ACTION ACT_ResetDrives:
// =============================================================
// ACT_ResetDrives
// Kasowanie bledow wszystkich falownikow
// =============================================================
//
// Dziala na ZBOCZE bitu xCmdResetDrives. Blok napedu wystawia
// impuls 200 ms na bicie 7 ControlWord - falownik NORD kasuje
// blad zboczem, nie poziomem.
//
// Kasujemy WSZYSTKIE napedy, takze te zablokowane w
// axDriveEnabled: skasowanie bledu niczego nie uruchamia,
// a chcemy widziec czysty obraz maszyny.
//
// Bit zdejmujemy sami, zeby nie trzeba bylo tego robic recznie
// w podgladzie online.

// -------------------------------------------------------------
// KASOWANIE RECZNE - bitem
// -------------------------------------------------------------

rtrgResetDrv(CLK := xCmdResetDrives);

IF rtrgResetDrv.Q THEN

	FOR i := 1 TO cNumDrives DO
		fbNord[i].M_Reset();
	END_FOR

	xCmdResetDrives	:= FALSE;
	xResetFailed	:= FALSE;

END_IF


// -------------------------------------------------------------
// KASOWANIE AUTOMATYCZNE - po wcisnieciu START
// -------------------------------------------------------------
//
// Kasujemy tylko te napedy, ktore faktycznie zglaszaja blad,
// i tylko ograniczona liczbe razy. Bez tego limitu maszyna
// dobijalaby sie w nieskonczonosc do napedu, ktory ma realny
// powod stac - a to wygladaloby jak "nic sie nie dzieje".

IF NOT xResetInProgress THEN
	RETURN;
END_IF


// Czysto - konczymy
IF NOT xAnyDriveFault THEN
	xResetInProgress	:= FALSE;
	nResetTries			:= 0;
	tonResetGap(IN := FALSE);
	RETURN;
END_IF


// Proby wyczerpane - dalej decyduje czlowiek
IF nResetTries >= cResetTries THEN
	xResetInProgress	:= FALSE;
	xResetFailed		:= TRUE;
	tonResetGap(IN := FALSE);
	RETURN;
END_IF


// Pierwsza proba od razu, kolejne co tResetGap
IF nResetTries = 0 THEN
	xDoResetPulse := TRUE;
ELSE
	tonResetGap(IN := TRUE, PT := tResetGap);
	xDoResetPulse := tonResetGap.Q;
END_IF

IF NOT xDoResetPulse THEN
	RETURN;
END_IF

tonResetGap(IN := FALSE);


FOR i := 1 TO cNumDrives DO
	IF axDrvFault[i] THEN
		fbNord[i].M_Reset();
	END_IF
END_FOR

nResetTries := nResetTries + 1;
END_ACTION

ACTION ACT_Sequence:
// =============================================================
// ACT_Sequence
// Wirtualna paleta idaca trasa maszyny
// =============================================================
//
// Paleta ZATRZYMUJE SIE na kazdej stacji. Cykl wyglada tak:
//
//   przejazd  para transporterow pracuje przez tStepTime,
//             potem OBA staja
//   praca     transportery stoja, dziala mechanika stacji
//             (kazdy ruch silownika przez tCylTime)
//   i dalej
//
// Czujnikow nie ma, wiec o zakonczeniu kazdej fazy decyduje
// czas. Po dolozeniu czujnikow te czasowki zastapi warunek
// "paleta na pozycji" i "silownik w polozeniu".
//
// TRASA:
//   poz. 1..11   dobre:   1-2-3-4-5-6-7-8-11-12-13
//   poz. 12..16  odrzut:  8-10-14-15-16  (8 -> 10 lancuchem)
//
// Przydzial falownikow do stacji:
//   st.1  -> 8     st.5  -> 5     st.9  -> 7      st.13 -> 15
//   st.2  -> 9     st.6  -> 6     st.10 -> 16     st.14 -> 17
//   st.3  -> 10    st.7  -> 11    st.11 -> 13     st.15 -> 18
//   st.4  -> 4     st.8  -> 12    st.12 -> 14     st.16 -> 19


// Zadanie ruchu kasujemy w kazdym cyklu - faza ustawia je od nowa
FOR i := 1 TO 20 DO
	axRunReq[i] := FALSE;
END_FOR

tThisStep := tCylTime;


// -------------------------------------------------------------
// START I STOP
// -------------------------------------------------------------

rtrgStart(CLK := START_TEST);

IF rtrgStart.Q THEN

	nIdx	:= 0;			// najpierw sprowadzamy mechanike
	nSub	:= 0;
	xMoving	:= FALSE;
	tonStep(IN := FALSE);

	xResetFailed := FALSE;
	nResetTries  := 0;
	tonResetGap(IN := FALSE);

	IF xAutoResetOnStart AND xAnyDriveFault THEN
		xResetInProgress := TRUE;
	END_IF

END_IF


IF NOT START_TEST THEN
	tonStep(IN := FALSE);
	sPhase := 'STOP - START_TEST = FALSE';
	ACT_ClearCoils();
	RETURN;
END_IF


IF NOT xSafetyOK THEN
	tonStep(IN := FALSE);
	sPhase := 'STOP - brak zezwolenia bezpieczenstwa';
	RETURN;
END_IF


IF xResetInProgress THEN
	tonStep(IN := FALSE);
	sPhase := CONCAT('kasowanie bledow falownikow - proba ',
	                 INT_TO_STRING(nResetTries));
	RETURN;
END_IF


// -------------------------------------------------------------
// TRYB RECZNY POJEDYNCZEGO SILOWNIKA
// -------------------------------------------------------------
//
// Ma pierwszenstwo przed sekwencja - transportery stoja,
// bo axRunReq zostalo wykasowane na gorze.

IF nManCyl <> 0 THEN
	ACT_ManualCyl();
	tonStep(IN := FALSE);
	RETURN;
END_IF


// -------------------------------------------------------------
// ZMIANA KROKU
// -------------------------------------------------------------
//
// Kazdy krok dostaje czasowke od zera i wlasne uzbrojenie
// czujnika. Bez tego krok dziedziczylby resztke po poprzednim.

xNewStep := (nIdx <> nIdxOld) OR (nSub <> nSubOld) OR (xMoving <> xMovingOld);

nIdxOld		:= nIdx;
nSubOld		:= nSub;
xMovingOld	:= xMoving;

IF xNewStep THEN
	tonStep(IN := FALSE);
	xStepArmed   := FALSE;
	xStepTimeout := FALSE;
END_IF


// Krok sam zglosi, na co czeka. Kasujemy co cykl.
xWaitSensor := FALSE;
xSensorOK   := FALSE;


// -------------------------------------------------------------
// FAZA
// -------------------------------------------------------------

IF xMoving THEN
	ACT_Move();
ELSE
	ACT_Work();
END_IF


// -------------------------------------------------------------
// KONIEC KROKU: CZUJNIK ALBO WATCHDOG
// -------------------------------------------------------------
//
// Krok czujnikowy konczy sie czujnikiem. Czasowka pracuje wtedy
// tylko jako watchdog - jesli to ONA zdecyduje, zapala sie
// xStepTimeout i wiadomo, ze czujnik nie przyszedl.
//
// Czujnik musi byc najpierw WOLNY (xStepArmed). Inaczej krok
// zaliczylby stan sprzed przejazdu albo czujnik zwarty na stale.

IF xUseSensors AND xWaitSensor THEN
	tThisStep := tMoveTimeout;
END_IF

tonStep(IN := TRUE, PT := tThisStep);
xAdvance := tonStep.Q;

// Watchdog wylaczony - czasowka nie ma prawa zakonczyc kroku
// czujnikowego. Krok stoi, dopoki nie przyjdzie sam czujnik.
IF xUseSensors AND xWaitSensor AND NOT xStepWatchdog THEN
	xAdvance := FALSE;
END_IF

IF xUseSensors AND xWaitSensor AND xAdvance THEN
	xStepTimeout := TRUE;
	nTimeouts    := nTimeouts + 1;
END_IF

IF NOT xSensorOK THEN
	xStepArmed := TRUE;
END_IF

IF xUseSensors AND xWaitSensor AND xStepArmed AND xSensorOK THEN
	xAdvance := TRUE;
END_IF

IF xAdvance THEN
	tonStep(IN := FALSE);
END_IF
END_ACTION

ACTION ACT_TestFeed:
// =============================================================
// ACT_TestFeed
// Proba calosciowa: st.1 -> desztaplarka -> stacja 4
// =============================================================
//
// Waska sciezka transportu na czas proby. NIE korzysta z tabeli
// trasy w ACT_Sequence - wozi tylko tam, gdzie trzeba:
//
//   1. dowozi stos ze stacji 1 na stacje 3 (czujnik IN2),
//   2. czeka, az desztaplarka zwolni palete,
//   3. wywozi ja przez stacje 4 robiac test dociskow,
//   4. ZATRZYMUJE ja na koncu stacji 4 - do recznego zabrania.
//
// Napedy: st.1 -> 8, st.2 -> 9, st.3 -> 10, st.4 -> 4.
// Rolki dociskowe (falownik 3) zostaja wylaczone.
//
// Cewki dociskow przepisujemy CO CYKL - ACT_ClearCoils zeruje
// je przy zdjetym START_TEST, wiec krok, ktory ich nie odswieza,
// stracilby sterowanie zaworem.


xFeedNewStep := (nFeedStep <> nFeedStepOld);
nFeedStepOld := nFeedStep;

IF xFeedNewStep THEN
	tonFeedStep(IN := FALSE);
	xFeedArmed := FALSE;
END_IF

tonFeedStep(IN := TRUE, PT := tFeedStep);
xFeedAdvance := tonFeedStep.Q AND NOT xFeedNewStep;


// Tor B ma WLASNA czasowke i wlasne uzbrojenie czujnika -
// inaczej dwie palety deptalyby sobie po jednym liczniku.
//
// UWAGA NA ZBOCZE KROKU MIEDZY TORAMI.
// Flagi xOutNewStep / xOutAdvance sa liczone TU, na poczatku
// akcji. Jesli inny tor wpisze torowi B numer kroku PO tym
// miejscu, krok wykona sie jeszcze w tym samym cyklu - ze stara
// flaga xOutAdvance, odziedziczona po kroku 0, gdzie czasowka
// dawno wybila. Krok przeskoczylby natychmiast.
//
// Wlasnie tak ginal przejazd ze stacji 5 na 6: krok 180 trwal
// JEDEN CYKL zadania, naped 5 dostawal zadanie na 10 ms i tor
// szedl dalej, jakby paleta juz przejechala.
//
// Dlatego zaden tor nie wpisuje numeru kroku innemu torowi.
// Zglasza tylko zadanie (xOutStart), a tor podnosi je SAM,
// w swoim kroku 0 - i wtedy pierwszy cykl nowego kroku jest
// juz zwyklym zboczem, z wyzerowana czasowka.

xOutNewStep := (nOutStep <> nOutStepOld);
nOutStepOld := nOutStep;

IF xOutNewStep THEN
	tonOutStep(IN := FALSE);
	xOutArmed := FALSE;
END_IF

tonOutStep(IN := TRUE, PT := tOutStep);
xOutAdvance := tonOutStep.Q AND NOT xOutNewStep;


xOut2NewStep := (nOut2Step <> nOut2StepOld);
nOut2StepOld := nOut2Step;

IF xOut2NewStep THEN
	tonOut2Step(IN := FALSE);
	xOut2Armed := FALSE;
END_IF

tonOut2Step(IN := TRUE, PT := tOut2Step);
xOut2Advance := tonOut2Step.Q AND NOT xOut2NewStep;


xOut3NewStep := (nOut3Step <> nOut3StepOld);
nOut3StepOld := nOut3Step;

IF xOut3NewStep THEN
	tonOut3Step(IN := FALSE);
	xOut3Armed := FALSE;
END_IF

tonOut3Step(IN := TRUE, PT := tOut3Step);
xOut3Advance := tonOut3Step.Q AND NOT xOut3NewStep;


// Czas pchania palety do blokady stacji 5 - liczony od wejscia
// w krok 80, niezalezny od czasowki kroku.
tonSt05Push(IN := (nFeedStep = 80), PT := tSt05_Push);

// Ile blokada stacji 5 stoi juz OPUSZCZONA. Nie ma na niej
// czujnika, wiec liczymy od zdjecia komendy wysuwu - tyle, ile
// dajemy kazdemu silownikowi na dojscie do polozenia.
tonSt05BlockDown(IN := NOT xFeed05_Block, PT := tCylTime);

// Od IN7 na stacji 8 do opuszczenia rolek pod paleta NOK.
// Liczona OSOBNO od tFeedSt08Stop - to sa dwie rozne rzeczy,
// wiec MOGA byc w dowolnej kolejnosci i dowolnie dalekie.
//
// Odliczamy od FLAGI OBECNOSCI, a nie od numeru kroku. Krok 215
// trwa tylko tFeedSt08Stop; przy dluzszym tSt08_DropDelay timer
// nie zdazyl dobiec do konca i zerowal sie przy przejsciu do
// kroku 218. Rolki nie schodzily wcale, a to, ze pierwsza paleta
// wygladala dobrze, robil krok 220 toru B3 - i tylko wtedy, gdy
// lancuch byl akurat wolny.
tonSt08Drop(IN := xSt08_AtStation, PT := tSt08_DropDelay);


rtrgFeedStart(CLK := START_FEED);

IF rtrgFeedStart.Q THEN
	nFeedStep  := 0;

	// Tor B tez od zera - inaczej po ponownym starcie dokanczal
	// by trase palety, ktorej juz tam nie ma.
	nOutStep   := 0;
	nOut2Step  := 0;
	nOut3Step  := 0;
	xSt05_Done := FALSE;
	xOutStart  := FALSE;
	xOut2Start := FALSE;
	xOut3Start := FALSE;
	xSt08_RollDown  := FALSE;
	xSt08_AtStation := FALSE;
END_IF


// Falowniki po zatrzymaniu runtime'u zglaszaja blad komunikacji
// i same z niego nie wyjda. Kasujemy go przy starcie, tak samo
// jak robi to START_TEST - inaczej za kazdym razem trzeba by
// pamietac o xCmdResetDrives.
IF rtrgFeedStart.Q AND xAutoResetOnStart AND xAnyDriveFault THEN
	xResetInProgress := TRUE;
	nResetTries      := 0;
	xResetFailed     := FALSE;
END_IF


// Domyslnie: cala mechanika w polozeniu spoczynkowym.
// Krok, ktory czegos potrzebuje, podaje to sam.
xFeedPressOn   := FALSE;
xFeedPressLoOn := FALSE;
xFeed05_Block  := FALSE;
xFeed05_Lift   := FALSE;
xFeed05_Jaws   := FALSE;
xFeed05_Pull   := FALSE;
tFeedStep      := tSt04_EntryToPress;
tOutStep       := tCylTime;
tOut2Step      := tCylTime;
tOut3Step      := tCylTime;

// Rolki domyslnie W GORZE - transport wzdluz. Tylko przejazd
// lancuchem opuszcza je swiadomie.
xFeedRoll08Up  := TRUE;
xFeedRoll10Up  := TRUE;


IF NOT START_FEED THEN
	sFeedPhase := 'DOWOZ - stop, START_FEED = FALSE';
END_IF


IF START_FEED AND xSafetyOK THEN

	CASE nFeedStep OF

	0:
		sFeedPhase := 'DOWOZ 0 czekam na potwierdzenie palet na st.1';

		// Bit SAM sie zdejmuje po przyjeciu. Dzieki temu po
		// oproznieniu stosu maszyna nie rusza w pustke, tylko
		// czeka na kolejne potwierdzenie operatora.
		//
		// Jesli IN2 juz widzi stos, to on STOI na stacji 3
		// i nie ma czego dowozic - idziemy od razu do pracy
		// desztaplarki. "Juz u celu" nie jest powodem do
		// czekania.
		IF xSt01_StackReady AND NOT xPal_St03 THEN
			xSt01_StackReady := FALSE;
			nFeedStep        := 10;
		END_IF

		IF xSt01_StackReady AND xPal_St03 THEN
			sFeedPhase       := 'DOWOZ 0 stos JUZ na st.3 - pomijam dowoz';
			xSt01_StackReady := FALSE;
			nFeedStep        := 20;
		END_IF

	10:
		sFeedPhase := 'DOWOZ 1 stos jedzie st.1 -> st.3, czekam na IN2';
		axRunReq[8]  := TRUE;
		axRunReq[9]  := TRUE;
		axRunReq[10] := TRUE;

		IF NOT xPal_St03 THEN xFeedArmed := TRUE; END_IF

		IF xPal_St03 AND NOT xFeedArmed THEN
			sFeedPhase := 'DOWOZ 1 IN2 JUZ zaslonony - odslon i zaslon ponownie';
		END_IF

		IF xFeedArmed AND xPal_St03 THEN nFeedStep := 15; END_IF

	15:
		// Dobieg po czujniku - stos dojezdza pod szczeki.
		// Przy tFeedSt03Stop = 0 krok trwa jeden cykl zadania.
		sFeedPhase := 'DOWOZ 1b dobieg stosu po IN2';
		axRunReq[9]  := TRUE;
		axRunReq[10] := TRUE;
		tFeedStep    := tFeedSt03Stop;

		IF xFeedAdvance THEN nFeedStep := 20; END_IF

	20:
		// Transportery STOJA - desztaplarka pracuje na stosie.
		sFeedPhase := 'DOWOZ 2 stos na st.3 - czekam na zwolnienie palety';

		IF xDe_PalletReleased THEN nFeedStep := 30; END_IF

	30:
		sFeedPhase := 'DOWOZ 3 paleta jedzie na st.4, czekam na IN3';

		// Paleta zaslaniajaca JUZ czujnik konca stacji 4 minela
		// wjazd pod rolki. Czekanie na IN3 bylo by czekaniem na
		// zdarzenie, ktore sie nie powtorzy - jedziemy dalej.
		IF xFeedNewStep AND xPal_St04End THEN
			sFeedPhase := 'DOWOZ 3 paleta JUZ na koncu st.4 - pomijam docisk';
			nFeedStep  := 75;
		END_IF

		axRunReq[10] := TRUE;
		axRunReq[4]  := TRUE;

		IF NOT xPal_St04In THEN xFeedArmed := TRUE; END_IF

		IF xPal_St04In AND NOT xFeedArmed THEN
			sFeedPhase := 'DOWOZ 3 IN3 JUZ zaslonony - odslon i zaslon ponownie';
		END_IF

		IF xFeedArmed AND xPal_St04In THEN nFeedStep := 40; END_IF

	40:
		sFeedPhase := 'ST.4 wjazd pod rolki - odstep przed dociskiem';
		axRunReq[10] := TRUE;
		axRunReq[4]  := TRUE;
		axRunReq[3]  := TRUE;   // rolki dociskowe
		tFeedStep    := tSt04_EntryToPress;

		IF xFeedAdvance THEN nFeedStep := 50; END_IF

	50:
		sFeedPhase := 'ST.4 dociski gorne schodza na deski';
		axRunReq[10] := TRUE;
		axRunReq[4]  := TRUE;
		axRunReq[3]  := TRUE;   // rolki dociskowe
		xFeedPressOn := TRUE;
		tFeedStep    := tSt04_UpToLo;

		IF xFeedAdvance THEN nFeedStep := 60; END_IF

	60:
		sFeedPhase := 'ST.4 TEST - czekam na koniec testu (IN4)';
		axRunReq[10]   := TRUE;
		axRunReq[4]    := TRUE;
		axRunReq[3]  := TRUE;   // rolki dociskowe
		xFeedPressOn   := TRUE;
		xFeedPressLoOn := TRUE;

		IF NOT xPal_St04End THEN xFeedArmed := TRUE; END_IF

		IF xPal_St04End AND NOT xFeedArmed THEN
			sFeedPhase := 'ST.4 IN4 JUZ zaslonony - odslon i zaslon ponownie';
		END_IF

		IF xFeedArmed AND xPal_St04End THEN nFeedStep := 70; END_IF

	70:
		// Dociski juz cofniete - kroki wyzej ich nie podaja.
		sFeedPhase := 'ST.4 koniec testu - dociski cofniete, dojazd';
		axRunReq[4] := TRUE;
		tFeedStep   := tSt04_StopDelay;

		IF xFeedAdvance THEN nFeedStep := 75; END_IF

	75:
		// BRAMKA MIEDZY TORAMI. Stacja 5 to zasob wspolny:
		// jej transporter i blokada obsluguja raz palete
		// wyjezdzajaca, raz wjezdzajaca. Wjazd moze ruszyc
		// dopiero wtedy, gdy poprzednia paleta zjechala ze
		// stacji 5 - czyli tor B jest wolny (0) albo minal
		// juz przejazd na stacje 6 (>= 200).
		//
		// Paleta czeka na koncu stacji 4, napedy stoja.
		sFeedPhase := 'ST.4 koniec - czekam, az zwolni sie stacja 5';

		IF (nOutStep = 0) OR (nOutStep >= 200) THEN
			nFeedStep := 80;
		END_IF

	80:
		// Blokada wysuwa sie RAZEM z ruszeniem palety ze stacji 4.
		// To ona zatrzymuje palete na stacji 5 - nie ma tam
		// czujnika, wiec musi czekac na palete, a nie odwrotnie.
		// Napedy pracuja TYLKO przez tSt05_Push, a nie przez caly
		// krok. Paleta opiera sie o blokade po kilku sekundach
		// i od tej chwili transporter mieli pod stojaca paleta -
		// tak przeciazylismy naped 5. Reszta kroku to juz tylko
		// uspokojenie palety, z zatrzymanymi napedami.
		sFeedPhase := 'ST.4 -> ST.5 przejazd, blokada juz wysunieta';
		xFeed05_Block := TRUE;
		tFeedStep   := tFeedToSt05;

		IF NOT tonSt05Push.Q THEN
			axRunReq[4] := TRUE;
			axRunReq[5] := TRUE;
		END_IF

		IF tonSt05Push.Q THEN
			sFeedPhase := 'ST.5 paleta na blokadzie - napedy staja';
		END_IF

		IF xFeedAdvance THEN nFeedStep := 100; END_IF


	// -----------------------------------------------------
	// STACJA 5 - TEST ROZRYWANIA
	// -----------------------------------------------------
	//
	// Transportery STOJA. Kolejnosc wg zalozen: blokada,
	// podniesienie szczek, chwyt, szesc silownikow rozrywajacych
	// w gore i w dol, zwolnienie, opuszczenie blokady.
	//
	// Kazdy krok podaje SWOJ pelny stan cewek - przepisujemy je
	// na dole akcji, w kazdym cyklu.

	100:
		// Paleta oparla sie o blokade. Transportery juz stoja,
		// dajemy jej uspokoic sie, zanim ruszy mechanika.
		sFeedPhase := 'ST.5 1/8 paleta na blokadzie - uspokojenie';
		xFeed05_Block := TRUE;
		tFeedStep     := tSt05_Settle;
		IF xFeedAdvance THEN nFeedStep := 110; END_IF

	110:
		sFeedPhase := 'ST.5 2/8 szczeki ida w gore';
		xFeed05_Block := TRUE;
		xFeed05_Lift  := TRUE;
		tFeedStep     := tCylTime;
		IF xFeedAdvance THEN nFeedStep := 120; END_IF

	120:
		sFeedPhase := 'ST.5 3/8 szczeki zamykaja sie na deskach';
		xFeed05_Block := TRUE;
		xFeed05_Lift  := TRUE;
		xFeed05_Jaws  := TRUE;
		tFeedStep     := tCylTime;
		IF xFeedAdvance THEN nFeedStep := 130; END_IF

	130:
		sFeedPhase := 'ST.5 4/8 ROZRYWANIE - silowniki ida w gore';
		xFeed05_Block := TRUE;
		xFeed05_Lift  := TRUE;
		xFeed05_Jaws  := TRUE;
		xFeed05_Pull  := TRUE;
		tFeedStep     := tCylTime;
		IF xFeedAdvance THEN nFeedStep := 140; END_IF

	140:
		sFeedPhase := 'ST.5 5/8 silowniki rozrywajace ida w dol';
		xFeed05_Block := TRUE;
		xFeed05_Lift  := TRUE;
		xFeed05_Jaws  := TRUE;
		tFeedStep     := tCylTime;
		IF xFeedAdvance THEN nFeedStep := 150; END_IF

	150:
		sFeedPhase := 'ST.5 6/8 szczeki otwieraja sie';
		xFeed05_Block := TRUE;
		xFeed05_Lift  := TRUE;
		tFeedStep     := tCylTime;
		IF xFeedAdvance THEN nFeedStep := 160; END_IF

	160:
		sFeedPhase := 'ST.5 7/8 szczeki ida w dol';
		xFeed05_Block := TRUE;
		tFeedStep     := tCylTime;
		IF xFeedAdvance THEN nFeedStep := 170; END_IF

	170:
		// PRZEKAZANIE PALETY TOROWI B.
		//
		// Tu konczy sie zadanie toru A. Paleta ma wolna droge
		// (blokada opuszczona) i od tej chwili jedzie na stacje
		// 16 SAMA, sekwencja nOutStep. Tor A wraca po nastepna.
		//
		// xSt05_Done to sygnal dla desztaplarki - na nim wydaje
		// kolejna palete, nie czekajac na stacje 16.
		//
		// Jesli tor B jeszcze pracuje, paleta czeka tutaj:
		// stoi na stacji 5 z opuszczona blokada, napedy staja.
		sFeedPhase := 'ST.5 8/8 blokada opuszcza sie';
		tFeedStep := tCylTime;

		// Oddajemy palete tylko wtedy, gdy tor B1 jest wolny
		// I stacja 7 pusta. Inaczej paleta zatrzymalaby sie
		// gdzies miedzy 5 a 6 i czekala tam bez potrzeby.
		xSt05_CanPass := (nOutStep = 0) AND NOT xPal_St07;

		IF xFeedAdvance AND NOT xSt05_CanPass THEN
			sFeedPhase := 'ST.5 gotowa - czekam, az zwolni sie droga na st.7';
		END_IF

		IF xFeedAdvance AND xSt05_CanPass AND (GVL_PERSIST.St03.Mem.nRemaining > 0) THEN
			nFeedPallets := nFeedPallets + 1;
			xOutStart    := TRUE;
			xSt05_Done   := TRUE;
			nFeedStep    := 20;
		END_IF

		IF xFeedAdvance AND xSt05_CanPass AND (GVL_PERSIST.St03.Mem.nRemaining <= 0) THEN
			nFeedPallets := nFeedPallets + 1;
			xOutStart    := TRUE;
			xSt05_Done   := TRUE;
			nFeedStep    := 0;
		END_IF

	END_CASE

END_IF


// =============================================================
// TOR B - STACJA 5 -> 16
// =============================================================
//
// Osobna sekwencja, wlasna czasowka (tOutStep / xOutAdvance)
// i wlasne uzbrojenie czujnika (xOutArmed). Startuje ja tor A
// w kroku 170, konczy sie zwolnieniem toru: nOutStep := 0.
//
// Czujniki mamy tylko na stacjach 7 (IN5), 8 (IN7) i 16
// (IN10). Reszta odcinkow konczy sie czasowka - kazda ma
// wlasna nazwe, zeby dalo sie ja dobrac osobno.
//
// Napedy toru B (5, 6, 11, 12, 7, 16..19) nie sa uzywane
// przez tor A - jedynym zasobem wspolnym jest naped 5
// i blokada stacji 5, rozdzielone bramka w kroku 75.

IF NOT START_FEED THEN
	sOutPhase := 'TOR B - stop, START_FEED = FALSE';
END_IF

IF START_FEED AND xSafetyOK THEN

	CASE nOutStep OF

	0:
		sOutPhase := 'TOR B wolny - czekam na palete ze stacji 5';

		IF xOutStart THEN
			xOutStart := FALSE;
			nOutStep  := 180;
		END_IF

	180:
		sOutPhase := 'ST.5 -> ST.6 przejazd';

		// Napedy i tak nie rusza, dopoki blokada nie opadnie -
		// pilnuje tego warunek nadrzedny w ACT_ApplyDrives.
		IF xSt05_BlockLock THEN
			sOutPhase := 'ST.5 czekam na opuszczenie blokady';
		END_IF

		axRunReq[5] := TRUE;
		axRunReq[6] := TRUE;
		tOutStep   := tFeed5to6;
		IF xOutAdvance THEN nOutStep := 200; END_IF

	200:
		// NIE WOLNO JECHAC W ZAJETE MIEJSCE.
		//
		// Dopoki czujnik jest zaslonony, a my nie jestesmy jeszcze
		// uzbrojeni, stoi tam CUDZA paleta - napedy musza stac.
		// Bez tego warunku transporter pchal palete w te, ktora
		// czekala na stacji 7, az do zderzenia; przy okazji
		// wykladalo to falownik stacji 5.
		sOutPhase := 'ST.6 -> ST.7 przejazd, czekam na IN5';

		// Przy 12 s w kroku 180 paleta potrafi dojechac na stacje 7
		// jeszcze przed wejsciem w ten krok. Stacja 7 byla pusta
		// w chwili przekazania (xSt05_CanPass), wiec zasloniety
		// czujnik NA WEJSCIU w krok to NASZA paleta - jest u celu,
		// nie ma na co czekac.
		IF xOutNewStep AND xPal_St07 THEN
			sOutPhase  := 'ST.7 paleta juz dojechala w kroku 180';
			nOutStep   := 205;
		END_IF

		IF NOT xPal_St07 OR xOutArmed THEN
			axRunReq[6]  := TRUE;
			axRunReq[11] := TRUE;
		END_IF

		IF NOT xPal_St07 THEN xOutArmed := TRUE; END_IF

		IF xPal_St07 AND NOT xOutArmed THEN
			sOutPhase := 'ST.7 ZAJETA - stoje, czekam az sie zwolni';
		END_IF

		IF xOutArmed AND xPal_St07 THEN nOutStep := 205; END_IF

	205:
		// Paleta LEZY na stacji 7, napedy staja. Tor B1 zwalnia
		// sie dopiero, gdy odbierze ja tor B2 - transporter
		// stacji 7 jest wspolny, wiec ruszajac nim po nastepna
		// palete pchnelibysmy te, ktora tu stoi.
		sOutPhase := 'ST.7 paleta czeka - tor B2 zajety';

		IF (nOut2Step = 0) AND ((nOut3Step = 0) OR (nOut3Step >= 240)) THEN
			sOutPhase  := 'ST.7 oddaje palete torowi B2';
			xOut2Start := TRUE;
			nOutStep   := 0;
		END_IF

	END_CASE

END_IF


// =============================================================
// TOR B2 - STACJA 7 -> STACJA 8
// =============================================================
//
// Krotki odcinek miedzy dwoma czujnikami: IN5 (st.7) i IN7
// (st.8). Wydzielony osobno, bo to on decyduje, kiedy stacja 7
// sie zwalnia i moze przyjac nastepna palete.
//
// Ruszy dopiero, gdy stacja 8 jest pusta - czyli tor B3 wolny.

IF START_FEED AND xSafetyOK THEN

	CASE nOut2Step OF

	0:
		sOut2Phase := 'TOR B2 wolny - stacja 7 moze oddac palete';

		IF xOut2Start THEN
			xOut2Start := FALSE;
			nOut2Step  := 210;
		END_IF

	210:
		// Jak w kroku 200: zaslonony czujnik przy nieuzbrojonym
		// kroku znaczy CUDZA paleta na stacji 8 - stoimy.
		sOut2Phase := 'ST.7 -> ST.8 przejazd, czekam na IN7';

		IF NOT xPal_St08 OR xOut2Armed THEN
			axRunReq[11] := TRUE;
			axRunReq[12] := TRUE;
		END_IF

		IF NOT xPal_St08 THEN xOut2Armed := TRUE; END_IF

		IF xPal_St08 AND NOT xOut2Armed THEN
			sOut2Phase := 'ST.8 ZAJETA - stoje, czekam az sie zwolni';
		END_IF

		IF xOut2Armed AND xPal_St08 THEN nOut2Step := 215; END_IF

	215:
		// Dobieg po IN7 - paleta dojezdza na srodek stacji 8,
		// zeby rolki mialy pod nia zejsc, a lancuch ja zabral.
		sOut2Phase := 'ST.8 dobieg po IN7';
		axRunReq[11] := TRUE;
		axRunReq[12] := TRUE;
		tOut2Step    := tFeedSt08Stop;

		// IN7 potwierdzone - paleta jest na stacji 8. Od tej chwili
		// biegnie odliczanie do opuszczenia rolek, niezaleznie od
		// tego, jak dlugo trwa ten krok i co bedzie dalej.
		xSt08_AtStation := TRUE;

		IF xOut2Advance THEN nOut2Step := 218; END_IF

	218:
		// Paleta stoi na srodku stacji 8, napedy staja. Czekamy,
		// az tor B3 sie zwolni - dopiero wtedy rolki moga zejsc
		// i lancuch ja zabrac.
		sOut2Phase := 'ST.8 paleta czeka - tor B3 zajety';

		IF nOut3Step = 0 THEN
			sOut2Phase := 'ST.8 oddaje palete torowi B3';
			xOut3Start := TRUE;
			nOut2Step  := 0;
		END_IF

	END_CASE

END_IF


// =============================================================
// TOR B3 - STACJA 8 -> LANCUCH -> 10 -> 14 -> 15 -> 16
// =============================================================
//
// Najdluzszy odcinek, bez czujnikow posrednich. Dopoki nim
// jedzie paleta, stacja 8 jest zajeta i tor B2 nie rusza.

IF START_FEED AND xSafetyOK THEN

	CASE nOut3Step OF

	0:
		sOut3Phase := 'TOR B3 wolny - stacja 8 moze oddac palete';

		IF xOut3Start THEN
			xOut3Start := FALSE;
			nOut3Step  := 220;
		END_IF

	220:
		// Paleta ma lec na lancuchu, wiec rolki OBU stacji schodza.
		sOut3Phase := 'ST.8 rolki 8 i 10 ida w dol - droga dla lancucha';
		xFeedRoll08Up := FALSE;
		xFeedRoll10Up := FALSE;
		tOut3Step     := tCylTime;
		IF xOut3Advance THEN nOut3Step := 230; END_IF

	230:
		// Jedzie SAM lancuch. Blokada w ACT_ApplyDrives i tak nie
		// pozwoli rolkom 8 i 10 ruszyc razem z falownikiem 7.
		sOut3Phase := 'ST.9 lancuch st.8 -> st.10';
		xFeedRoll08Up := FALSE;
		xFeedRoll10Up := FALSE;
		axRunReq[7]   := TRUE;
		tOut3Step     := tFeed9Chain;
		IF xOut3Advance THEN nOut3Step := 240; END_IF

	240:
		sOut3Phase := 'ST.10 rolki ida w gore - paleta jedzie na 14';
		tOut3Step := tCylTime;
		IF xOut3Advance THEN nOut3Step := 250; END_IF

	250:
		sOut3Phase := 'ST.10 -> ST.14 przejazd';
		axRunReq[16] := TRUE;
		axRunReq[17] := TRUE;
		tOut3Step    := tFeed10to14;
		IF xOut3Advance THEN nOut3Step := 260; END_IF

	260:
		sOut3Phase := 'ST.14 -> ST.15 przejazd';
		axRunReq[17] := TRUE;
		axRunReq[18] := TRUE;
		tOut3Step    := tFeed14to15;
		IF xOut3Advance THEN nOut3Step := 270; END_IF

	270:
		// Jak wyzej: na stacji 16 moze jeszcze lezec paleta,
		// ktorej operator nie odebral. Nie wpychamy w nia kolejnej.
		sOut3Phase := 'ST.15 -> ST.16 przejazd, czekam na IN10';

		IF NOT xPal_St16 OR xOut3Armed THEN
			axRunReq[18] := TRUE;
			axRunReq[19] := TRUE;
		END_IF

		IF NOT xPal_St16 THEN xOut3Armed := TRUE; END_IF

		IF xPal_St16 AND NOT xOut3Armed THEN
			sOut3Phase := 'ST.16 ZAJETA - stoje, czekam az operator odbierze';
		END_IF

		IF xOut3Armed AND xPal_St16 THEN
			nFeedPallets := nFeedPallets + 1;
			nOut3Step    := 275;
		END_IF

	275:
		sOut3Phase := 'ST.16 dobieg po IN10';
		axRunReq[18] := TRUE;
		axRunReq[19] := TRUE;
		tOut3Step    := tFeedSt16Stop;

		IF xOut3Advance THEN nOut3Step := 280; END_IF

	280:
		// Paleta stoi na stacji 16. Odbiera ja operator - gdy
		// zniknie z czujnika, po tSt16_Clear tor B sie zwalnia
		// i moze przyjac nastepna palete ze stacji 5.
		//
		// Tor B NIE decyduje juz, czy jechac po nastepna palete
		// - to nalezy do toru A i desztaplarki.
		sOut3Phase := 'ST.16 paleta odebrana - czekam na oproznienie';
		tOut3Step  := tSt16_Clear;

		IF xPal_St16 THEN
			sOut3Phase := 'ST.16 paleta STOI - odbierz ja';
			tonOut3Step(IN := FALSE);
		END_IF

		IF NOT xPal_St16 AND xOut3Advance THEN
			nOut3Step := 0;
		END_IF

	END_CASE

END_IF


// =============================================================
// ROLKI STACJI 8 W DOLE - ZATRZASK
// =============================================================
//
// Raz opuszczone pod paleta NOK rolki maja tam zostac, az
// lancuch przewiezie palete na stacje 10. Inaczej kazdy krok,
// ktory ich nie pisze, podniosl by je z powrotem i paleta
// podskakiwalaby miedzy rolkami a lancuchem.
//
// Zatrzask zdejmujemy NA ZBOCZU wejscia w krok 240 toru B3,
// czyli w chwili, gdy lancuch dowiozl palete na stacje 10.
//
// MUSI to byc zbocze, nie poziom. Warunek poziomowy
// (nOut3Step >= 240) jest prawdziwy przez CALA dalsza trase
// az do stacji 16 - a ta regula wykonuje sie PO krokach.
// Nastepna paleta zapalala wiec zatrzask w kroku 215, a ten
// warunek gasil go w tym samym cyklu. Rolki schodzily dopiero
// wtedy, gdy operator zabral palete ze stacji 16 i tor B3
// wrocil do zera. Tak to wygladalo na maszynie: pierwsza
// paleta dobrze, kazda nastepna duzo za pozno.
//
// Rolek stacji 10 to NIE dotyczy - nimi steruje tor B3.

IF xOut3NewStep AND (nOut3Step = 240) THEN
	xSt08_RollDown  := FALSE;
	xSt08_AtStation := FALSE;
END_IF

// DRUGIE KASOWANIE - siatka bezpieczenstwa.
//
// Wjazd nastepnej palety na stacje 8 (krok 210 toru B2) wymaga
// rolek W GORZE. Gdyby zatrzask z jakiegokolwiek powodu przezyl
// poprzednia palete, nastepna nie mialaby po czym wjechac i
// staloby to tak dlugo, az ktos zabierze palete z konca linii.
//
// W tym momencie poprzedniej palety nad rolkami juz nie ma -
// tor B2 nie ruszylby, gdyby stacja 8 byla zajeta.

IF xOut2NewStep AND (nOut2Step = 210) THEN
	xSt08_RollDown  := FALSE;
	xSt08_AtStation := FALSE;
END_IF

// Opuszczenie rolek. Warunek nadrzedny, nie krok - paleta ma
// siasc na lancuchu tSt08_DropDelay po IN7, obojetne czy tor B2
// jest jeszcze w dobiegu, czy juz czeka na zwolnienie lancucha.

IF xSt08_PalletNOK AND xSt08_AtStation AND tonSt08Drop.Q THEN
	xSt08_RollDown := TRUE;
END_IF

IF xSt08_RollDown THEN
	xFeedRoll08Up := FALSE;
END_IF


// =============================================================
// CZY ZADANE NAPEDY MOGA RUSZYC
// =============================================================
//
// Krok mowi, czego oczekuje od czujnikow. Ale jesli naped nie
// moze ruszyc, paleta nigdy nie dojedzie i fraza o czujniku
// jest mylaca - wyglada, jakby zawinil czujnik.
//
// Szukamy PIERWSZEGO zadanego napedu, ktory nie potwierdza
// pracy, i nazywamy przyczyne od skutku do zrodla: pozniejsze
// przypisanie wygrywa, wiec zostaje przyczyna najglebsza.

nFeedBadDrv := 0;
sFeedDrvWhy := '';

// Przyczyne ustalamy W PETLI, po indeksie i - nigdy po
// nFeedBadDrv, ktore moze byc zerem. ST nie gwarantuje
// skrocenia obliczen w AND, wiec zapis axDrvFault[nFeedBadDrv]
// siegalby poza tablice ARRAY[1..20] przy braku zadan.

FOR i := 1 TO cNumDrives DO

	IF axRunReq[i] AND NOT axDrvRunning[i] AND (nFeedBadDrv = 0) THEN

		nFeedBadDrv := i;
		sFeedDrvWhy := 'nie potwierdza pracy';

		IF axDrvFault[i] THEN
			sFeedDrvWhy := 'BLAD - kasuj xCmdResetDrives';
		END_IF

		IF NOT axDriveEnabled[i] THEN
			sFeedDrvWhy := 'NIEDOPUSZCZONY w axDriveEnabled';
		END_IF

	END_IF

END_FOR


// Chwilowy brak potwierdzenia to normalny rozbieg, dopiero
// utrzymujacy sie jest problemem.
tonFeedDrv(IN := START_FEED AND (nFeedBadDrv > 0), PT := T#2S);

IF START_FEED AND tonFeedDrv.Q THEN
	sFeedPhase := CONCAT('NAPED ', INT_TO_STRING(nFeedBadDrv));
	sFeedPhase := CONCAT(sFeedPhase, ' STOI: ');
	sFeedPhase := CONCAT(sFeedPhase, sFeedDrvWhy);
END_IF


// -------------------------------------------------------------
// DOCISKI STACJI 4 -> CEWKI, CO CYKL
// -------------------------------------------------------------
//
// Gorne schodza pierwsze, dolne po tSt04_UpToLo, cofaja sie
// razem. Przepisujemy w kazdym cyklu, zeby nic nie moglo
// zabrac sterowania zaworem w trakcie jazdy.

IF START_FEED THEN
	xSt04_UpExt := xFeedPressOn;
	xSt04_UpRet := NOT xFeedPressOn;
	xSt04_LoExt := xFeedPressLoOn;
	xSt04_LoRet := NOT xFeedPressLoOn;
END_IF


// -------------------------------------------------------------
// ROLKI PODNOSZONE 8 i 10 -> CEWKI, CO CYKL
// -------------------------------------------------------------

IF START_FEED THEN
	xSt08_Up   := xFeedRoll08Up;
	xSt08_Down := NOT xFeedRoll08Up;
	xSt10_Up   := xFeedRoll10Up;
	xSt10_Down := NOT xFeedRoll10Up;
END_IF


// -------------------------------------------------------------
// MECHANIKA STACJI 5 -> CEWKI, CO CYKL
// -------------------------------------------------------------

IF START_FEED THEN

	xSt05_BlockExt := xFeed05_Block;
	xSt05_BlockRet := NOT xFeed05_Block;

	xSt05_LiftUp   := xFeed05_Lift;
	xSt05_LiftDown := NOT xFeed05_Lift;

	xSt05_JawClose := xFeed05_Jaws;

	FOR i := 1 TO 6 DO
		axSt05_PullUp[i]   := xFeed05_Pull;
		axSt05_PullDown[i] := NOT xFeed05_Pull;
	END_FOR

END_IF
END_ACTION

ACTION ACT_Work:
// =============================================================
// ACT_Work
// Praca stacji - transportery STOJA
// =============================================================
//
// Kazdy ruch silownika trwa tCylTime. Stacje bez mechaniki
// przechodza od razu do przejazdu.

CASE nIdx OF


// -------------------------------------------------------------
// 0 - SPROWADZENIE MECHANIKI DO POLOZENIA WYJSCIOWEGO
// -------------------------------------------------------------

0:
	sPhase := 'polozenie wyjsciowe mechaniki';

	xSt03_JawClose := FALSE;
			xSt03_JawOpen  := TRUE;
	xSt11_JawClose := FALSE;
			xSt11_JawOpen  := TRUE;

	xSt04_UpExt := FALSE;	xSt04_UpRet := TRUE;
	xSt04_LoExt := FALSE;	xSt04_LoRet := TRUE;

	xSt05_BlockExt := FALSE;
			xSt05_BlockRet := TRUE;
	xSt05_LiftUp   := FALSE;
			xSt05_LiftDown := TRUE;
	xSt05_JawClose := FALSE;
	FOR i := 1 TO 6 DO
				axSt05_PullUp[i]   := FALSE;
				axSt05_PullDown[i] := TRUE;
			END_FOR

	xSt08_Up   := TRUE;
	xSt08_Down := FALSE;
	xSt10_Up   := TRUE;
	xSt10_Down := FALSE;

	IF xAdvance THEN
		nIdx	:= 1;
		nSub	:= 0;
		xMoving	:= FALSE;
	END_IF


// -------------------------------------------------------------
// 1 - STACJA 1: CZEKAMY NA STOS
// -------------------------------------------------------------
//
// Czujnika IN1 nie uzywamy. Jedziemy dopiero, gdy operator
// (albo pozniej czujnik) postawi xSt01_StackReady na TRUE.
// Krok nie ma czasowki - stoi, dopoki bit nie przyjdzie.

1:
	sPhase := 'st.1 czekam na stos - bit xSt01_StackReady';

	IF xSt01_StackReady THEN
		sPhase := 'st.1 stos gotowy - jazda';
		xMoving	:= TRUE;
		nSub	:= 0;
	END_IF


// -------------------------------------------------------------
// 3 - DESZTAPLARKA: SAME SZCZEKI
// -------------------------------------------------------------
//
// Wozek stoi - falownik 1 jest zablokowany, mechanika
// podnoszenia niegotowa. Sprawdzamy tylko zawory szczek.

3:
	CASE nSub OF
		0:
			sPhase := 'st.3 szczeki zamykaja sie';
			xSt03_JawClose := TRUE;
			xSt03_JawOpen  := FALSE;
			IF xAdvance THEN nSub := 10; END_IF
		10:
			sPhase := 'st.3 szczeki otwieraja sie';
			xSt03_JawClose := FALSE;
			xSt03_JawOpen  := TRUE;
			IF xAdvance THEN xMoving := TRUE; nSub := 0; END_IF
	END_CASE


// -------------------------------------------------------------
// 4 - KONIEC TESTU SCISKANIA
// -------------------------------------------------------------
//
// Sam test odbyl sie na JADACEJ palecie, w ACT_MoveSt04. Tutaj
// paleta juz stoi na koncu stacji, a my tylko pilnujemy, zeby
// dociski byly cofniete, zanim ruszy dalej.

4:
	sPhase := 'st.4 test zakonczony - dociski cofniete';
	xSt04_UpExt := FALSE;	xSt04_UpRet := TRUE;
	xSt04_LoExt := FALSE;	xSt04_LoRet := TRUE;
	IF xAdvance THEN xMoving := TRUE; nSub := 0; END_IF


// -------------------------------------------------------------
// 5 - TEST ROZRYWANIA
// -------------------------------------------------------------

5:
	CASE nSub OF
		0:
			sPhase := 'st.5 blokada wysuwa sie';
			xSt05_BlockExt := TRUE;
			xSt05_BlockRet := FALSE;
			IF xAdvance THEN nSub := 10; END_IF
		10:
			sPhase := 'st.5 szczeki ida w gore';
			xSt05_LiftUp   := TRUE;
			xSt05_LiftDown := FALSE;
			IF xAdvance THEN nSub := 20; END_IF
		20:
			sPhase := 'st.5 szczeki zamykaja sie';
			xSt05_JawClose := TRUE;
			IF xAdvance THEN nSub := 30; END_IF
		30:
			sPhase := 'st.5 silowniki rozrywajace ida w gore';
			FOR i := 1 TO 6 DO
				axSt05_PullUp[i]   := TRUE;
				axSt05_PullDown[i] := FALSE;
			END_FOR
			IF xAdvance THEN nSub := 40; END_IF
		40:
			sPhase := 'st.5 silowniki rozrywajace ida w dol';
			FOR i := 1 TO 6 DO
				axSt05_PullUp[i]   := FALSE;
				axSt05_PullDown[i] := TRUE;
			END_FOR
			IF xAdvance THEN nSub := 50; END_IF
		50:
			sPhase := 'st.5 szczeki otwieraja sie';
			xSt05_JawClose := FALSE;
			IF xAdvance THEN nSub := 60; END_IF
		60:
			sPhase := 'st.5 szczeki ida w dol';
			xSt05_LiftUp   := FALSE;
			xSt05_LiftDown := TRUE;
			IF xAdvance THEN nSub := 70; END_IF
		70:
			sPhase := 'st.5 blokada opuszcza sie';
			xSt05_BlockExt := FALSE;
			xSt05_BlockRet := TRUE;
			IF xAdvance THEN xMoving := TRUE; nSub := 0; END_IF
	END_CASE


// -------------------------------------------------------------
// 8 - ROZJAZD, PRZEBIEG DOBRYCH: ROLKI W GORZE
// -------------------------------------------------------------

8:
	sPhase := 'st.8 rolki ida w gore - paleta jedzie prosto';
	xSt08_Up   := TRUE;
	xSt08_Down := FALSE;
	IF xAdvance THEN xMoving := TRUE; nSub := 0; END_IF


// -------------------------------------------------------------
// 9 - SZTAPLARKA: SAME SZCZEKI
// -------------------------------------------------------------

9:
	CASE nSub OF
		0:
			sPhase := 'st.11 szczeki zamykaja sie';
			xSt11_JawClose := TRUE;
			xSt11_JawOpen  := FALSE;
			IF xAdvance THEN nSub := 10; END_IF
		10:
			sPhase := 'st.11 szczeki otwieraja sie';
			xSt11_JawClose := FALSE;
			xSt11_JawOpen  := TRUE;
			IF xAdvance THEN xMoving := TRUE; nSub := 0; END_IF
	END_CASE


// -------------------------------------------------------------
// 11 - WYJSCIE DOBRYCH, KONIEC PRZEBIEGU
// -------------------------------------------------------------

11:
	sPhase := 'st.13 odbior - nowa paleta na stacji 8, trasa odrzutu';
	IF xAdvance THEN
		nIdx	:= 12;
		nSub	:= 0;
		xMoving	:= FALSE;
	END_IF


// -------------------------------------------------------------
// 12 - ROZJAZD, PRZEBIEG ODRZUTU: OBIE ROLKI W DOLE
// -------------------------------------------------------------
//
// Paleta ma lezec na lancuchu, wiec rolki stacji 8 I 10 musza
// zejsc, zanim lancuch ruszy.

12:
	CASE nSub OF
		0:
			sPhase := 'st.8 rolki ida w dol';
			xSt08_Up   := FALSE;
	xSt08_Down := TRUE;
			IF xAdvance THEN nSub := 10; END_IF
		10:
			sPhase := 'st.10 rolki ida w dol - droga dla lancucha';
			xSt10_Up   := FALSE;
	xSt10_Down := TRUE;
			IF xAdvance THEN xMoving := TRUE; nSub := 0; END_IF
	END_CASE


// -------------------------------------------------------------
// 13 - PRZEKIEROWANIE: ROLKI W GORE
// -------------------------------------------------------------

13:
	sPhase := 'st.10 rolki ida w gore - paleta jedzie na 14';
	xSt10_Up   := TRUE;
	xSt10_Down := FALSE;
	IF xAdvance THEN xMoving := TRUE; nSub := 0; END_IF


// -------------------------------------------------------------
// 16 - ODBIOR ODRZUTU, KONIEC PETLI
// -------------------------------------------------------------

16:
	sPhase := 'st.16 odbior - koniec przebiegu';
	IF xAdvance THEN
		nIdx	:= 0;
		nSub	:= 0;
		xMoving	:= FALSE;
		nLoops	:= nLoops + 1;
	END_IF


// -------------------------------------------------------------
// STACJE BEZ MECHANIKI - postoj i jedziemy dalej
// -------------------------------------------------------------

ELSE
	sPhase := 'postoj na stacji - brak mechaniki';
	IF xAdvance THEN xMoving := TRUE; nSub := 0; END_IF

END_CASE
END_ACTION

END_PROGRAM

(* stored: Version 1.1.0.1
   POU MAIN: Id {3723006f-8e56-479b-b982-5b261f2b6738}, SpecialFunc None
   Action ACT_ApplyDrives: Id {4a10e003-0000-4000-9000-00000000e003}
   Action ACT_CamCycles: Id {4a10e011-0000-4000-9000-000000000011}
   Action ACT_ClearCoils: Id {4a10e009-0000-4000-9000-00000000e009}
   Action ACT_Config: Id {4a10e001-0000-4000-9000-00000000e001}
   Action ACT_Drives: Id {4a10e004-0000-4000-9000-00000000e004}
   Action ACT_Inputs: Id {4a10e00f-0000-4000-9000-00000000e00f}
   Action ACT_Logger: Id {4a10e013-0000-4000-9000-000000000013}
   Action ACT_LogRow: Id {4a10e014-0000-4000-9000-000000000014}
   Action ACT_ManualCyl: Id {4a10e00a-0000-4000-9000-00000000e00a}
   Action ACT_Move: Id {4a10e007-0000-4000-9000-00000000e007}
   Action ACT_MoveSt04: Id {4a10e010-0000-4000-9000-000000000010}
   Action ACT_Outputs: Id {4a10e008-0000-4000-9000-00000000e008}
   Action ACT_ResetDrives: Id {4a10e005-0000-4000-9000-00000000e005}
   Action ACT_Sequence: Id {4a10e002-0000-4000-9000-00000000e002}
   Action ACT_TestFeed: Id {4a10e012-0000-4000-9000-000000000012}
   Action ACT_Work: Id {4a10e006-0000-4000-9000-00000000e006} *)
